SUBAPPLICATION NumericValue_TO_AUI2_AND_STORE (* Wie MyLib::sys::NumericValue_TO_AUI2 (VT lesen, als bidirektionalen AUI2-Plug an einen Consumer wie AOption_AUI_DEMUX_N.K weiterreichen), zusaetzlich mit INI-Persistenz: beim Boot gewinnt der aus INI_AUI2 geladene Wert (per AUI_LAST_2 gegen die Live-VT-Lesung gemergt), danach jede Live-Aenderung; gespeichert wird immer der vom Consumer ZURUECKGEMELDETE (tatsaechlich uebernommene) Wert. Eigene Baustein-Klasse getrennt von INI_IN_AND_STORE_AUI2/ _AUDI2 - die bleiben unveraendert (KEY/SECTION, plain VALUEO), da sie in zahlreichen anderen Projekten verwendet werden. *)
  (* Standard: 61499-2; Description: Copyright (c) 2026 Meisterschulen am Ostbahnhof This program and the accompanying materials are made available under the terms of the Eclipse Public License 2.0 which is available at https://www.eclipse.org/legal/epl-2.0/ SPDX-License-Identifier: EPL-2.0 *)
  (* Version 3.1, 2026-11-13, Franz Höpfinger, Meisterschulen am Ostbahnhof, Neuer Eingang DEFAULT_VALUE (bisher fest 0) an INI_AUI.DEFAULT_VALUE - je Instanz einstellbar, Default unveraendert 0. *)
  (* Version 3.0, 2026-10-13, Franz Höpfinger, Meisterschulen am Ostbahnhof, Korrektur 2: der bisher ungenutzte Boot-Wert von INI_AUI2 (AUI_TO_AUI2_1.AUI_OUT) wird jetzt tatsaechlich verwendet - per AUI_LAST_2 (Last-Writer-Wins) gegen die Live-VT-Lesung (AD_TO_AUI.AUI_OUT) gemergt, bevor es zu VALUEO geht. Da SETM=FALSE ist, feuert INI_AUI2 dieses Boot-Echo nur einmal beim Start (INIT->INITO->GET->GETO), nicht bei jedem spaeteren Schreibvorgang - kein Dauerkreislauf. *)
  (* Version 2.0, 2026-10-13, Franz Höpfinger, Meisterschulen am Ostbahnhof, Korrektur: die Live-VT-Lesung geht jetzt DIREKT an VALUEO (ein einziges AUI_TO_AUI2, wie in NumericValue_TO_AUI2) - NICHT mehr ueber INI_AUI2 vorgeschaltet. Gespeichert wird stattdessen erst das vom Consumer ueber VALUEO ZURUECKGEMELDETE (tatsaechlich uebernommene) Ergebnis, ueber eine zweite, reine Schreib-Bruecke zu INI_AUI2. SETM=FALSE (statt TRUE) verhindert, dass INI_AUI2 jeden Schreibvorgang sofort wieder quittiert/zurueckmeldet - das wuerde sich sonst im Kreis drehen (Wert raus, zurueck, erneut speichern, erneut raus, ...), da dieses Echo hier nirgendwo terminiert wird. *)
  PACKAGE MyLib::sys;
  IMPORT isobus::UT::Q::const::IDs::ID_NULL;
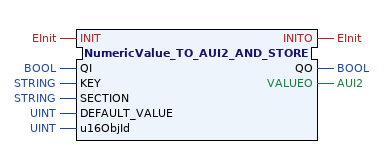
  EVENT_INPUT
    INIT : EInit; (* Initialization Request *)
  END_EVENT
  EVENT_OUTPUT
    INITO : EInit; (* Initialization Confirm *)
  END_EVENT
  VAR_INPUT
    QI : BOOL := TRUE; (* Quality Input - TRUE to enable service *)
    KEY : STRING; (* Key name. *)
    SECTION : STRING; (* Section name. *)
    DEFAULT_VALUE : UINT := UINT#0; (* Wert, wenn der KEY noch nicht in der INI steht *)
    u16ObjId : UINT := ID_NULL; (* Object ID *)
  END_VAR
  VAR_OUTPUT
    QO : BOOL; (* Quality Output - TRUE if service executed successfully *)
  END_VAR
  PLUGS
    VALUEO : adapter::types::bidirectional::AUI2;
  END_PLUGS
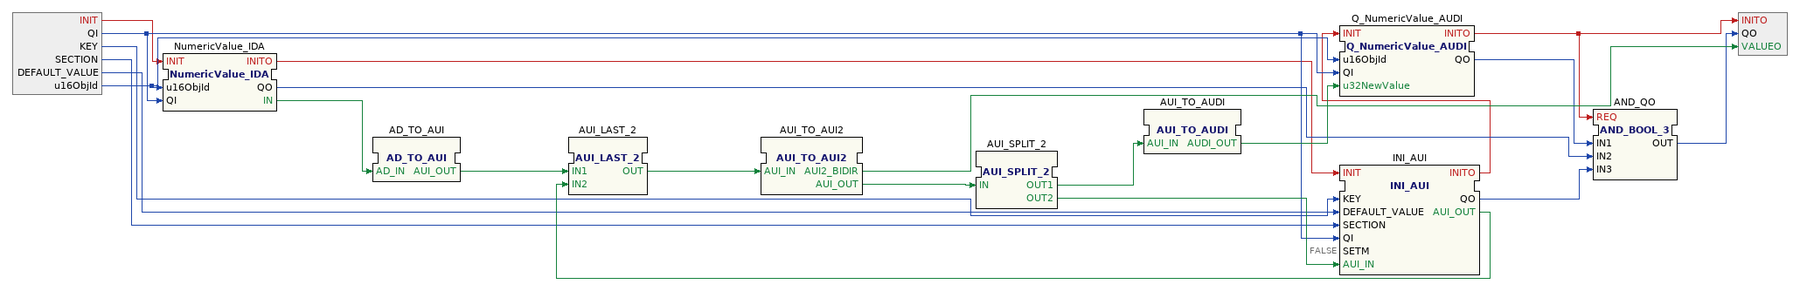
  (* SETM=FALSE: INI_AUI2 quittiert nur beim Boot (INIT->INITO->GET->GETO) automatisch, NICHT bei jedem spaeteren Schreibvorgang ueber VAL (Vorwaertsrichtung). Der Boot-Wert laeuft ueber AUI_TO_AUI2_1.AUI_OUT zu AUI_LAST_2 (siehe oben) und gewinnt dort einmalig gegen die Live-VT-Lesung. Waere SETM=TRUE, wuerde jeder spaetere Schreibvorgang sofort ein neues Echo auf AUI_OUT ausloesen, das wieder bei AUI_LAST_2 ankaeme und erneut Richtung VALUEO geschickt wuerde - ein Dauerkreislauf. *)
  FBS
    NumericValue_IDA : isobus::UT::io::NumericValue::NumericValue_IDA;
    AD_TO_AUI : adapter::conversion::unidirectional::AD_TO_AUI;
    AUI_TO_AUI2 : adapter::conversion::bidirectional::AUI_TO_AUI2; (* Bruecke zum externen Consumer (z.B. AOption_AUI_DEMUX_N.K) *)
    AUI_TO_AUDI : adapter::conversion::unidirectional::AUI_TO_AUDI;
    Q_NumericValue_AUDI : isobus::UT::Q::Q_NumericValue_AUDI;
    AUI_LAST_2 : adapter::events::unidirectional::AUI_LAST_2; (* Last-Writer-Wins: beim Boot gewinnt der INI_AUI2-Wert (IN2), danach jede Live-VT-Aenderung (IN1) *)
    AUI_SPLIT_2 : adapter::events::unidirectional::AUI_SPLIT_2;
    INI_AUI : eclipse4diac::storage::INI_AUI(SETM := FALSE);
    AND_QO : iec61131::booleanOperators::AND_BOOL_3;
  END_FBS
  EVENT_CONNECTIONS
    INIT TO NumericValue_IDA.INIT;
    NumericValue_IDA.INITO TO INI_AUI.INIT;
    INI_AUI.INITO TO Q_NumericValue_AUDI.INIT;
    Q_NumericValue_AUDI.INITO TO INITO;
    Q_NumericValue_AUDI.INITO TO AND_QO.REQ;
  END_CONNECTIONS
  DATA_CONNECTIONS
    KEY TO INI_AUI.KEY;
    DEFAULT_VALUE TO INI_AUI.DEFAULT_VALUE;
    SECTION TO INI_AUI.SECTION;
    u16ObjId TO NumericValue_IDA.u16ObjId;
    u16ObjId TO Q_NumericValue_AUDI.u16ObjId;
    QI TO Q_NumericValue_AUDI.QI;
    QI TO NumericValue_IDA.QI;
    QI TO INI_AUI.QI;
    Q_NumericValue_AUDI.QO TO AND_QO.IN1;
    NumericValue_IDA.QO TO AND_QO.IN2;
    INI_AUI.QO TO AND_QO.IN3;
    AND_QO.OUT TO QO;
  END_CONNECTIONS
  ADAPTER_CONNECTIONS
    NumericValue_IDA.IN TO AD_TO_AUI.AD_IN;
    AD_TO_AUI.AUI_OUT TO AUI_LAST_2.IN1;
    AUI_LAST_2.OUT TO AUI_TO_AUI2.AUI_IN;
    AUI_TO_AUI2.AUI2_BIDIR TO VALUEO;
    AUI_TO_AUDI.AUDI_OUT TO Q_NumericValue_AUDI.u32NewValue;
    AUI_SPLIT_2.OUT1 TO AUI_TO_AUDI.AUI_IN;
    AUI_SPLIT_2.OUT2 TO INI_AUI.AUI_IN;
    INI_AUI.AUI_OUT TO AUI_LAST_2.IN2;
    AUI_TO_AUI2.AUI_OUT TO AUI_SPLIT_2.IN;
  END_CONNECTIONS
END_SUBAPPLICATION
